(* IEC 61131-3 sources: krc-sample-programs/motor-ramp-alarms-codesys/source/08_Alarms, 4 files *)

(* ---- E_AlarmLevel.st ---- *)
// How serious an alarm is.
TYPE E_AlarmLevel :
(
	LVL_INFO    := 1,	// Shows on the alarm list. Nothing else
	LVL_WARNING := 2,	// Lights the orange light. The machine keeps running
	LVL_ALARM   := 3 	// Stops the machine: the state machine goes to Fault until it is cleared
) INT;
END_TYPE

(* ---- ST_Alarm.st ---- *)
// One line of the alarm table. The level and the text are filled in where the table is declared
// (GVL_Alarms). bTriggered is wired by one line per alarm in ALARMS; the rest belongs to the alarm
// list in ALARMS.
TYPE ST_Alarm :
STRUCT
	eLevel      : E_AlarmLevel;	// INFO, WARNING or ALARM (set in the table)
	sText       : STRING(60);	// What happened, in words, for the screen (set in the table)
	bTriggered  : BOOL;	// The condition, right now (ALARMS, one line per alarm)
	bOnList     : BOOL;	// On the list: from when it triggers until it is acknowledged and gone (ALARMS)
	bAcked      : BOOL;	// Acknowledged with ACK or Reset (ALARMS)
	iStepRaised : INT;	// The step the machine was in when it came on (ALARMS)
END_STRUCT
END_TYPE

(* ---- ST_Permissive.st ---- *)
// One line of the permissive table: something Ready waits for. The text is filled in where the table
// is declared (GVL_Alarms); bSatisfied is wired by one line per permissive in DEVICES.
TYPE ST_Permissive :
STRUCT
	sText       : STRING(30);	// What Ready waits for, in words (set in the table)
	bSatisfied  : BOOL;	// Met, right now (DEVICES, one line per permissive)
END_STRUCT
END_TYPE

(* ---- GVL_Alarms.st ---- *)
// The alarm table and the permissive table: every alarm and every permissive, with its words, in one
// place. Adding an alarm is a line here, a constant in CONSTANTS, and its trigger line in ALARMS.
VAR_GLOBAL
	aAlarms : ARRAY[1..ALARM_COUNT] OF ST_Alarm := [
		(eLevel := LVL_ALARM,   sText := 'E-stop pressed: the safety circuit is open'),
		(eLevel := LVL_ALARM,   sText := 'Drive dropped out while running'),
		(eLevel := LVL_ALARM,   sText := 'Drive switched to local while running'),
		(eLevel := LVL_ALARM,   sText := 'Ramp timeout: speed not reached in time'),
		(eLevel := LVL_ALARM,   sText := 'Stop timeout: the motor did not stop in time'),
		(eLevel := LVL_WARNING, sText := 'Speed deviation: more than 10 % off'),
		(eLevel := LVL_INFO,    sText := 'Simulation mode: SIM is playing the machine')];
	aPermissives : ARRAY[1..PERMISSIVE_COUNT] OF ST_Permissive := [
		(sText := 'Drive ready'),
		(sText := 'Drive in remote'),
		(sText := 'Stop released'),
		(sText := 'Motor stopped')];
	bAlarmOnList     : BOOL;	// Any ALARM-level alarm on the list (ALARMS)
	bWarningOnList   : BOOL;	// Any WARNING on the list (ALARMS)
	bUnacknowledged  : BOOL;	// Any ALARM or WARNING on the list not yet acknowledged (ALARMS)
	bPermissivesOK   : BOOL;	// Every permissive met (STATE_MACHINE)
END_VAR
